(* IEC 61131-3 sources: SemaPLC/sema-plc-benchmark/spec2control-benchmark/data/st-baseline/tennessee-eastman-chemical/pous/programs, 8 files *)

(* ---- main.st ---- *)
PROGRAM main
VAR
	Heartbeat : bool;
END_VAR

(* Entry point required by OpenPLC Editor v4. The process sections run as parallel program instances under task0; main only provides a scan heartbeat. *)
Heartbeat := NOT Heartbeat;

END_PROGRAM

(* ---- Section2.st ---- *)
PROGRAM Section2
VAR
	FIT101_Flow_PV_GPM : real;
	PI001_Pressure_PV_psig : real;
	FIC104_MV_to_PV103_Pct : real;
	FIT_101 : ANALOG_IN;
	PI_001 : ANALOG_IN;
	FIC_104 : PID_BASIC;
	PV_103 : VALVE_ELECTRIC;
	XV_106 : VALVE_ON_OFF;
	IAL_101 : BOOL_INPUT;
	FAL_101 : DIGITAL_IN;
	FAL_102 : DIGITAL_IN;
	FAL_103 : DIGITAL_IN;
	XV106NotOpen : bool;
	XV106Interlock : bool;
	FIC104Inhibit : bool;
END_VAR

FIT_101(
    PV_High := 180.0,
    PV_Low := 40.0,
    Scaling_Slope := 12.5,
    Scaling_Offset := -50.0,
    Alarm_Enable := TRUE);
PI_001(
    Alarm_Enable := TRUE);
FAL_101(
    DI_Raw := FIT_101.High_Alarm);
FAL_102(
    DI_Raw := FIT_101.Low_Alarm);
FAL_103(
    DI_Raw := FIT_101.General_Fault);
XV_106();
XV106NotOpen := NOT XV_106.FB_Opened;
XV106Interlock := XV106NotOpen OR XV_106.Alarm_Position_Error OR XV_106.Alarm_General;
IAL_101(
    Bool_In := XV106Interlock,
    Alarm_OnTrue := TRUE,
    Latch_Enable := TRUE);
FIC104Inhibit := IAL_101.Bool_Out OR FAL_103.DI_Out OR PI_001.High_Alarm OR PI_001.Low_Alarm;
FIC_104(
    PV := FIT_101.PV,
    SP := 100.0,
    MV_MIN := 0.0,
    MV_MAX := 100.0,
    X0 := 0.0,
    KP := 1.5,
    TR := 0.6,
    TD := 0.1,
    Inhibit := FIC104Inhibit);
PV_103(
    Control_Signal := FIC_104.XOUT,
    Manual_Position := 0.0,
    Open_Limit := 100.0,
    Close_Limit := 0.0,
    Inhibit := FAL_103.DI_Out);

(* Outputs published to other sections / HMI. *)
FIT101_Flow_PV_GPM := FIT_101.PV;
PI001_Pressure_PV_psig := PI_001.PV;
FIC104_MV_to_PV103_Pct := FIC_104.XOUT;

END_PROGRAM

(* ---- Section3.st ---- *)
PROGRAM Section3
VAR
	TIT_103_Temperature_C : real;
	LT_105_Level_Percent : real;
	TIC_101_Output_Percent : real;
	LIC_106_Output_Percent : real;
	TIT_103 : ANALOG_IN;
	LT_105 : ANALOG_IN;
	TIC_101 : PID_BASIC;
	LIC_106 : PID_BASIC;
	FC_004 : PID_BASIC;
	LV_104 : VALVE_ELECTRIC;
	XV_102 : VALVE_ON_OFF;
	TIC101_Inhibit_OR : bool;
	SteamNotOpen_NOT : bool;
	LIC106_Inhibit_OR : bool;
END_VAR

TIT_103(
    PV_High := 200.0,
    PV_Low := 160.0,
    Scaling_Slope := 15.625,
    Scaling_Offset := -62.5,
    Alarm_Enable := TRUE);
LT_105(
    PV_High := 80.0,
    PV_Low := 20.0,
    Scaling_Slope := 6.25,
    Scaling_Offset := -25.0,
    Alarm_Enable := TRUE);
FC_004();
XV_102(
    Timeout := T#5s,
    Inhibit := TIT_103.High_Alarm);
TIC101_Inhibit_OR := TIT_103.High_Alarm OR XV_102.Alarm_Position_Error OR FC_004.PV_Low_Alarm OR TIT_103.General_Fault;
TIC_101(
    PV := TIT_103.PV,
    SP := 180.0,
    MV_MIN := 0.0,
    MV_MAX := 100.0,
    KP := 3.0,
    TR := 1.2,
    TD := 0.1,
    Inhibit := TIC101_Inhibit_OR);
LV_104(
    Control_Signal := LIC_106.XOUT,
    Open_Limit := 100.0,
    Close_Limit := 0.0,
    Inhibit := LT_105.High_Alarm);
SteamNotOpen_NOT := NOT XV_102.FB_Opened;
LIC106_Inhibit_OR := SteamNotOpen_NOT OR LV_104.Alarm OR LT_105.General_Fault;
LIC_106(
    PV := LT_105.PV,
    SP := 50.0,
    MV_MIN := 0.0,
    MV_MAX := 100.0,
    KP := 2.5,
    TR := 0.9,
    TD := 0.0,
    Inhibit := LIC106_Inhibit_OR);

(* Outputs published to other sections / HMI. *)
TIT_103_Temperature_C := TIT_103.PV;
LT_105_Level_Percent := LT_105.PV;
TIC_101_Output_Percent := TIC_101.XOUT;
LIC_106_Output_Percent := LIC_106.XOUT;

END_PROGRAM

(* ---- Section4.st ---- *)
PROGRAM Section4
VAR
	FIT103_FlowRate : real;
	LT104_Level : real;
	LIC101_PV102_ValveCommand : real;
	LAH101_Alarm : bool;
	LAL101_Alarm : bool;
	LT104_FaultAlarm : bool;
	OverCapacity_Active : bool;
	LevelAbove10_OK : bool;
	FIT_103 : ANALOG_IN;
	LT_104 : ANALOG_IN;
	LIC_101 : PID_BASIC;
	PV_102 : VALVE_ELECTRIC;
	OverCapCompare : bool;
	SPOverrideSelector : real;
	LevelAbove10Compare : bool;
	LevelLowInvert : bool;
	PV102InhibitLogic : bool;
	LT104AutoInvert : bool;
END_VAR

FIT_103(
    Scaling_Slope := 3.125,
    Scaling_Offset := -12.5,
    Alarm_Enable := TRUE);
LT_104(
    Scaling_Slope := 6.25,
    Scaling_Offset := -25.0,
    Alarm_Enable := TRUE);
LT104AutoInvert := NOT LT_104.General_Fault;
OverCapCompare := (FIT_103.PV > 60.0);
SPOverrideSelector := SEL(G := OverCapCompare, IN0 := 65.0, IN1 := 50.0);
LIC_101(
    AUTO := LT104AutoInvert,
    PV := LT_104.PV,
    SP := SPOverrideSelector,
    MV_MIN := 0.0,
    MV_MAX := 100.0,
    X0 := 0.0,
    KP := 1.8,
    TR := 0.6,
    TD := 0.1,
    PV_High := 90.0,
    PV_Low := 15.0,
    Deviation_Limit := 5.0);
LevelAbove10Compare := (LT_104.PV > 10.0);
LevelLowInvert := NOT LevelAbove10Compare;
PV102InhibitLogic := LevelLowInvert OR LT_104.General_Fault;
PV_102(
    Control_Signal := LIC_101.XOUT,
    Manual_Mode := FALSE,
    Manual_Position := 0.0,
    Open_Limit := 100.0,
    Close_Limit := 0.0,
    Timeout := T#10s,
    Inhibit := PV102InhibitLogic);

(* Outputs published to other sections / HMI. *)
FIT103_FlowRate := FIT_103.PV;
LT104_Level := LT_104.PV;
LIC101_PV102_ValveCommand := LIC_101.XOUT;
LAH101_Alarm := LIC_101.PV_High_Alarm;
LAL101_Alarm := LIC_101.PV_Low_Alarm;
LT104_FaultAlarm := LT_104.General_Fault;
OverCapacity_Active := OverCapCompare;
LevelAbove10_OK := LevelAbove10Compare;

END_PROGRAM

(* ---- Section5.st ---- *)
PROGRAM Section5
VAR
	TIT106_ReboilerTemp_PV : real;
	LT107_Column2Level_PV : real;
	TIC106_FV105_SteamFlow_MV : real;
	LIC107_LV102_Outflow_MV : real;
	TIT_106 : ANALOG_IN;
	LT_107 : ANALOG_IN;
	TIC_106 : PID_BASIC;
	LIC_107 : PID_BASIC;
	FV_105 : VALVE_ELECTRIC;
	LV_102 : VALVE_ELECTRIC;
	CONDENSATE_RETURN_VALVE_OPEN_LS : DIGITAL_IN;
	SteamValveInhibitLogic : bool;
	CondensateNotOpen : bool;
END_VAR

TIT_106(
    PV_High := 260.0,
    Scaling_Slope := 18.75,
    Scaling_Offset := -75.0,
    Alarm_Enable := TRUE);
LT_107(
    PV_High := 80.0,
    PV_Low := 20.0,
    Scaling_Slope := 6.25,
    Scaling_Offset := -25.0,
    Alarm_Enable := TRUE);
TIC_106(
    AUTO := TRUE,
    PV := TIT_106.PV,
    SP := 200.0,
    MV_MIN := 0.0,
    MV_MAX := 100.0,
    KP := -3.0,
    TR := 1.2,
    TD := 0.2);
LIC_107(
    AUTO := TRUE,
    PV := LT_107.PV,
    SP := 50.0,
    MV_MIN := 0.0,
    MV_MAX := 100.0,
    KP := 2.5,
    TR := 1.0,
    TD := 0.0);
CONDENSATE_RETURN_VALVE_OPEN_LS();
CondensateNotOpen := NOT CONDENSATE_RETURN_VALVE_OPEN_LS.DI_Out;
SteamValveInhibitLogic := CondensateNotOpen OR TIC_106.PV_High_Alarm;
FV_105(
    Control_Signal := TIC_106.XOUT,
    Open_Limit := 100.0,
    Close_Limit := 0.0,
    Inhibit := SteamValveInhibitLogic);
LV_102(
    Control_Signal := LIC_107.XOUT,
    Open_Limit := 100.0,
    Close_Limit := 0.0,
    Inhibit := LIC_107.PV_Low_Alarm);

(* Outputs published to other sections / HMI. *)
TIT106_ReboilerTemp_PV := TIT_106.PV;
LT107_Column2Level_PV := LT_107.PV;
TIC106_FV105_SteamFlow_MV := TIC_106.XOUT;
LIC107_LV102_Outflow_MV := LIC_107.XOUT;

END_PROGRAM

(* ---- Section7.st ---- *)
PROGRAM Section7
VAR
	TI_008_Temp_PV : real;
	LI_003_Level_PV : real;
	TIC_106_MV_Pct : real;
	LIC_103_MV_Pct : real;
	XV_105_Valve_Position_Pct : real;
	XV_104_Valve_Position_Pct : real;
	Column3_Start_CMD : bool;
	TIC106_DeviationFault : bool;
	LIC101_Condensate_High : bool;
	LI_003 : ANALOG_IN;
	TI_008 : ANALOG_IN;
	LIC_103 : PID_BASIC;
	TIC_106 : PID_BASIC;
	XV_104 : VALVE_ELECTRIC;
	XV_105 : VALVE_ELECTRIC;
	LIC_101_HI : BOOL_INPUT;
	StartDelay_TON : TON;
	TIC106_DevTON : TON;
	TI8_GT_200 : bool;
	InhibitFinal_OR : bool;
	LI3_Above30_GT : bool;
	SteamStartPermissive_AND : bool;
	InhibitNot_NOT : bool;
	TIC106_Auto_AND : bool;
	LI3_Below15_GT : bool;
	XV104_Close_OR : bool;
	XV104_AutoNot_NOT : bool;
END_VAR

LI_003(
    PV_Low := 10.0,
    Scaling_Slope := 6.25,
    Scaling_Offset := -25.0,
    Alarm_Enable := TRUE);
TI_008(
    PV_High := 195.0,
    Scaling_Slope := 15.625,
    Scaling_Offset := -62.5,
    Alarm_Enable := TRUE);
LI3_Below15_GT := (15.0 > LI_003.PV);
XV104_Close_OR := LI_003.Low_Alarm OR LI3_Below15_GT;
XV104_AutoNot_NOT := NOT XV104_Close_OR;
LIC_103(
    AUTO := XV104_AutoNot_NOT,
    PV := LI_003.PV,
    SP := 70.0,
    MV_MIN := 0.0,
    MV_MAX := 100.0,
    KP := 2.5,
    TR := 0.8,
    TD := 0.1);
LIC_101_HI(
    Bool_In := LIC101_Condensate_High,
    Alarm_OnTrue := TRUE);
TI8_GT_200 := (TI_008.PV > 200.0);
InhibitFinal_OR := TI8_GT_200 OR LIC_101_HI.Bool_Out;
InhibitNot_NOT := NOT InhibitFinal_OR;
LI3_Above30_GT := (LI_003.PV > 30.0);
StartDelay_TON(
    IN := Column3_Start_CMD,
    PT := T#12s);
SteamStartPermissive_AND := StartDelay_TON.Q AND LI3_Above30_GT;
TIC106_Auto_AND := SteamStartPermissive_AND AND InhibitNot_NOT;
TIC_106(
    AUTO := TIC106_Auto_AND,
    PV := TI_008.PV,
    SP := 180.0,
    MV_MIN := 5.0,
    MV_MAX := 95.0,
    X0 := 0.0,
    KP := -3.2,
    TR := 1.0,
    TD := 0.3,
    Deviation_Limit := 10.0,
    Inhibit := InhibitFinal_OR);
XV_104(
    Control_Signal := LIC_103.XOUT,
    Manual_Mode := XV104_Close_OR,
    Manual_Position := 0.0,
    Open_Limit := 100.0,
    Close_Limit := 0.0,
    Timeout := T#10s);
XV_105(
    Control_Signal := TIC_106.XOUT,
    Open_Limit := 100.0,
    Close_Limit := 0.0,
    Timeout := T#10s,
    Inhibit := InhibitFinal_OR);
TIC106_DevTON(
    IN := TIC_106.Deviation_Alarm,
    PT := T#30s);

(* Outputs published to other sections / HMI. *)
TIC106_DeviationFault := TIC106_DevTON.Q;
TI_008_Temp_PV := TI_008.PV;
LI_003_Level_PV := LI_003.PV;
TIC_106_MV_Pct := TIC_106.XOUT;
LIC_103_MV_Pct := LIC_103.XOUT;
XV_105_Valve_Position_Pct := XV_105.Valve_Position;
XV_104_Valve_Position_Pct := XV_104.Valve_Position;

END_PROGRAM

(* ---- Section8.st ---- *)
PROGRAM Section8
VAR
	LT102_Level_PV_Pct : real;
	FIT105_Flow_PV_LPM : real;
	LIC106_MV_To_XV101_Pct : real;
	FC008_MV_To_PV104_Pct : real;
	Decanter2_Online : bool;
	FIT_105 : ANALOG_IN;
	LT_102 : ANALOG_IN;
	LT_103 : ANALOG_IN;
	LT_107 : ANALOG_IN;
	LIC_106 : PID_BASIC;
	FC_008 : PID_BASIC;
	XV_101 : VALVE_ELECTRIC;
	PV_104 : VALVE_ELECTRIC;
	LIC106_StartupDelay : TON;
	FC8_StartupDelay : TON;
	LT102_SignalFaults_A : bool;
	LT102_SignalFaults : bool;
	LT103_Above90Check : bool;
	LIC106_ForceClose_A : bool;
	LIC106_ForceClose : bool;
	LIC106_ForceCloseClear : bool;
	LIC106_AutoEnable : bool;
	FIT105_HighLow : bool;
	FIT105_Invalid : bool;
	FC8_SignalValid : bool;
	LT107_Below20Check : bool;
	FC8_NoForceClose : bool;
	FC8_AutoBase : bool;
	FC8_AutoInterlocks : bool;
	FC8_AutoEnable : bool;
	FC8_ForceOpen : bool;
	FC8_InhibitLogic : bool;
END_VAR

FIT_105(
    Scaling_Slope := 9.375,
    Scaling_Offset := -37.5,
    Alarm_Enable := TRUE);
LT_102(
    Scaling_Slope := 6.25,
    Scaling_Offset := -25.0,
    Alarm_Enable := TRUE);
LT_103(
    PV_High := 85.0,
    Scaling_Slope := 6.25,
    Scaling_Offset := -25.0,
    Alarm_Enable := TRUE);
LT_107(
    PV_Low := 15.0,
    Scaling_Slope := 6.25,
    Scaling_Offset := -25.0,
    Alarm_Enable := TRUE);
LT102_SignalFaults_A := LT_102.High_Alarm OR LT_102.Low_Alarm;
LT102_SignalFaults := LT102_SignalFaults_A OR LT_102.General_Fault;
LT103_Above90Check := (LT_103.PV > 90.0);
LIC106_ForceClose_A := LT103_Above90Check OR LT102_SignalFaults;
XV_101(
    Control_Signal := LIC_106.XOUT,
    Manual_Mode := LIC106_ForceClose,
    Manual_Position := 0.0,
    Timeout := T#10s,
    Inhibit := LIC106_ForceClose);
LIC106_ForceClose := LIC106_ForceClose_A OR XV_101.Alarm;
LIC106_ForceCloseClear := NOT LIC106_ForceClose;
LIC106_StartupDelay(
    IN := TRUE,
    PT := T#14s);
LIC106_AutoEnable := LIC106_StartupDelay.Q AND LIC106_ForceCloseClear;
LIC_106(
    AUTO := LIC106_AutoEnable,
    PV := LT_102.PV,
    SP := 65.0,
    MV_MIN := 0.0,
    MV_MAX := 100.0,
    X0 := 0.0,
    KP := -3.0,
    TR := 1.2,
    TD := 0.0,
    Inhibit := LIC106_ForceClose);
FIT105_HighLow := FIT_105.High_Alarm OR FIT_105.Low_Alarm;
FIT105_Invalid := FIT105_HighLow OR FIT_105.General_Fault;
FC8_SignalValid := NOT FIT105_Invalid;
FC8_StartupDelay(
    IN := TRUE,
    PT := T#14s);
FC8_AutoBase := FC8_StartupDelay.Q AND FC8_SignalValid;
LT107_Below20Check := (LT_107.PV < 20.0);
FC8_NoForceClose := NOT LT107_Below20Check;
FC8_AutoInterlocks := Decanter2_Online AND FC8_NoForceClose;
FC8_AutoEnable := FC8_AutoBase AND FC8_AutoInterlocks;
PV_104(
    Control_Signal := FC_008.XOUT,
    Manual_Mode := LT107_Below20Check,
    Manual_Position := 0.0,
    Inhibit := FC8_InhibitLogic);
FC8_ForceOpen := FIT_105.General_Fault OR PV_104.Alarm;
FC8_InhibitLogic := LT107_Below20Check OR FC8_ForceOpen;
FC_008(
    AUTO := FC8_AutoEnable,
    PV := FIT_105.PV,
    SP := 120.0,
    MV_MIN := 0.0,
    MV_MAX := 100.0,
    X0 := 100.0,
    KP := 2.5,
    TR := 0.8,
    TD := 0.2,
    Deviation_Limit := 12.0,
    Inhibit := FC8_InhibitLogic);

(* Outputs published to other sections / HMI. *)
LT102_Level_PV_Pct := LT_102.PV;
FIT105_Flow_PV_LPM := FIT_105.PV;
LIC106_MV_To_XV101_Pct := LIC_106.XOUT;
FC008_MV_To_PV104_Pct := FC_008.XOUT;

END_PROGRAM

(* ---- Section9.st ---- *)
PROGRAM Section9
VAR
	TIT101_Temperature_PV_C : real;
	FI103_Flow_PV : real;
	FIC103_Output_MV_Percent : real;
	LV102_ValvePositionCmd_Percent : real;
	XV104_Open_FB : bool;
	LC002_ValidLevel : bool;
	LC002_LevelValid_In : bool;
	TIT_101 : ANALOG_IN;
	FI_103 : ANALOG_IN;
	FIC_103 : PID_BASIC;
	LV_102 : VALVE_ELECTRIC;
	XV_104 : VALVE_ON_OFF;
	LC_002 : BOOL_INPUT;
	XV104NotOpen_NOT : bool;
	LC002NotActive_NOT : bool;
	LV102Inhibit_OR : bool;
	XV104Inhibit_OR : bool;
	FIC103Inhibit_OR : bool;
	XV104OpenCmd_NOT : bool;
END_VAR

TIT_101(
    PV_High := 55.0,
    Scaling_Slope := 6.25,
    Scaling_Offset := -25.0,
    Alarm_Enable := TRUE);
FI_103(
    PV_Low := 5.0,
    Scaling_Slope := 6.25,
    Scaling_Offset := -25.0,
    Alarm_Enable := TRUE);
LC_002(
    Bool_In := LC002_LevelValid_In);
LC002NotActive_NOT := NOT LC_002.Bool_Out;
FIC103Inhibit_OR := TIT_101.General_Fault OR TIT_101.Low_Alarm OR LC002NotActive_NOT;
FIC_103(
    AUTO := TRUE,
    PV := TIT_101.PV,
    SP := 45.0,
    MV_MIN := 0.0,
    MV_MAX := 100.0,
    X0 := 0.0,
    KP := 3.0,
    TR := 1.2,
    TD := 0.3,
    Inhibit := FIC103Inhibit_OR);
XV104Inhibit_OR := FI_103.Low_Alarm OR TIT_101.High_Alarm;
XV104OpenCmd_NOT := NOT XV104Inhibit_OR;
XV_104(
    Open_Cmd := XV104OpenCmd_NOT,
    Close_Cmd := XV104Inhibit_OR,
    Timeout := T#2s,
    Inhibit := XV104Inhibit_OR);
XV104NotOpen_NOT := NOT XV_104.FB_Opened;
LV102Inhibit_OR := XV104NotOpen_NOT OR FI_103.Low_Alarm OR TIT_101.General_Fault OR LC002NotActive_NOT OR TIT_101.High_Alarm OR XV_104.Alarm_General;
LV_102(
    Control_Signal := FIC_103.XOUT,
    Manual_Mode := FALSE,
    Manual_Position := 0.0,
    Open_Limit := 100.0,
    Close_Limit := 0.0,
    Timeout := T#2s,
    Inhibit := LV102Inhibit_OR);

(* Outputs published to other sections / HMI. *)
TIT101_Temperature_PV_C := TIT_101.PV;
FI103_Flow_PV := FI_103.PV;
FIC103_Output_MV_Percent := FIC_103.XOUT;
LV102_ValvePositionCmd_Percent := LV_102.Valve_Position;
XV104_Open_FB := XV_104.FB_Opened;
LC002_ValidLevel := LC_002.Bool_Out;

END_PROGRAM
